// Model of the TwinSAFE FB SR (set dominant latch).
// The Safety Editor refuses an SR with Set or Reset unconnected: the model then reports Error with
// diagnostic bit 15 instead of running (see T_SafeFunctionBlockBase).
{attribute 'reflection'}
FUNCTION_BLOCK T_SafeSr EXTENDS T_SafeFunctionBlockBase
VAR_INPUT
    Set : BOOL;
    Reset : BOOL;
    Parameters : ST_SafeLatchParameters;
END_VAR
VAR_OUTPUT
    SrOut : BOOL;
END_VAR
VAR
    {attribute 'is_connected' := 'Set'}
    _setConnected : BOOL;
    {attribute 'is_connected' := 'Reset'}
    _resetConnected : BOOL;
    _state : E_SafeLatchState := E_SafeLatchState.Stop;
END_VAR

SUPER^();

// Set and Reset must both be connected (Safety Editor: "Inport Set of SR must be connected").
METHOD PROTECTED ConfigurationOk : BOOL
IF NOT _setConnected THEN
    _configurationFault := 'T_SafeSr: Inport Set of SR must be connected';
    RETURN;
ELSIF NOT _resetConnected THEN
    _configurationFault := 'T_SafeSr: Inport Reset of SR must be connected';
    RETURN;
END_IF

ConfigurationOk := TRUE;
END_METHOD

METHOD PROTECTED Process
VAR
    setActive : BOOL;
    resetActive : BOOL;
END_VAR
setActive   := F_SafeInputValue(_setConnected, Parameters.SetMakeContact, Set);
resetActive := F_SafeInputValue(_resetConnected, Parameters.ResetMakeContact, Reset);

IF NOT _fbRun THEN
    _state := E_SafeLatchState.Stop;
ELSE
    IF _state = E_SafeLatchState.Stop THEN
        _state := E_SafeLatchState.Safe;
    END_IF

    IF setActive THEN
        _state := E_SafeLatchState.Set;
    ELSIF resetActive THEN
        _state := E_SafeLatchState.Safe;
    END_IF
END_IF

SrOut := (_state = E_SafeLatchState.Set);
Error := FALSE;
Diag  := 0;
State := TO_BYTE(_state);
END_METHOD

END_FUNCTION_BLOCK

(* stored: Version 1.1.0.1
   POU T_SafeSr: Id {f012fcb5-00f3-58d8-85cf-893035478446}, SpecialFunc None
   Method ConfigurationOk: Id {15455a7b-ca7d-4dbc-a1fd-6d40b3e632d8}
   Method Process: Id {7e42194a-8cb8-5273-8753-b28131026d06} *)
